Staubli VAL3: cycle_Hold.pgx

program cycle_Hold()
begin
  //cycle进程:Holding
  rs:_nOmacStat=5
  //if isPowered()
  //    disablePower()
  //    watch(isPowered()==false,2)
  //  endIf
  stopMove()
  wait(isSettled())
  //cycle进程:Held
  rs:_nOmacStat=6
  logMsg("当前处于暂停状态 "+toString(".2",clock()))
  rs:_sRobotStatus="当前处于暂停状态"
end
